FUNCTION_BLOCK CASE_SEQUENCER (* Solvability control: ecc_persistent form, designed by hand. Never shown to a model. *)
  (* Standard: 61499-2 *)
  (* Version 1.0, 2026-11-06, st2fb *)
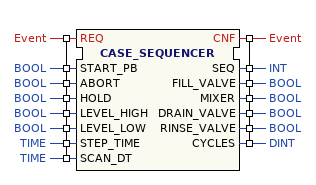
  EVENT_INPUT
    REQ WITH START_PB, ABORT, HOLD, LEVEL_HIGH, LEVEL_LOW, STEP_TIME, SCAN_DT;
  END_EVENT
  EVENT_OUTPUT
    CNF WITH SEQ, FILL_VALVE, MIXER, DRAIN_VALVE, RINSE_VALVE, CYCLES;
  END_EVENT
  VAR_INPUT
    START_PB : BOOL;
    ABORT : BOOL;
    HOLD : BOOL;
    LEVEL_HIGH : BOOL;
    LEVEL_LOW : BOOL;
    STEP_TIME : TIME;
    SCAN_DT : TIME;
  END_VAR
  VAR_OUTPUT
    SEQ : INT;
    FILL_VALVE : BOOL;
    MIXER : BOOL;
    DRAIN_VALVE : BOOL;
    RINSE_VALVE : BOOL;
    CYCLES : DINT;
  END_VAR
  VAR
    TIMING : BOOL;
    ST2FB_NOW : TIME;
    STEP_TIMER_IN : BOOL;
    STEP_TIMER_PT : TIME;
    STEP_TIMER_Q : BOOL;
    STEP_TIMER_ET : TIME;
    STEP_TIMER_STATE : INT;
    STEP_TIMER_PREV_IN : BOOL;
    STEP_TIMER_START_TIME : TIME;
  END_VAR
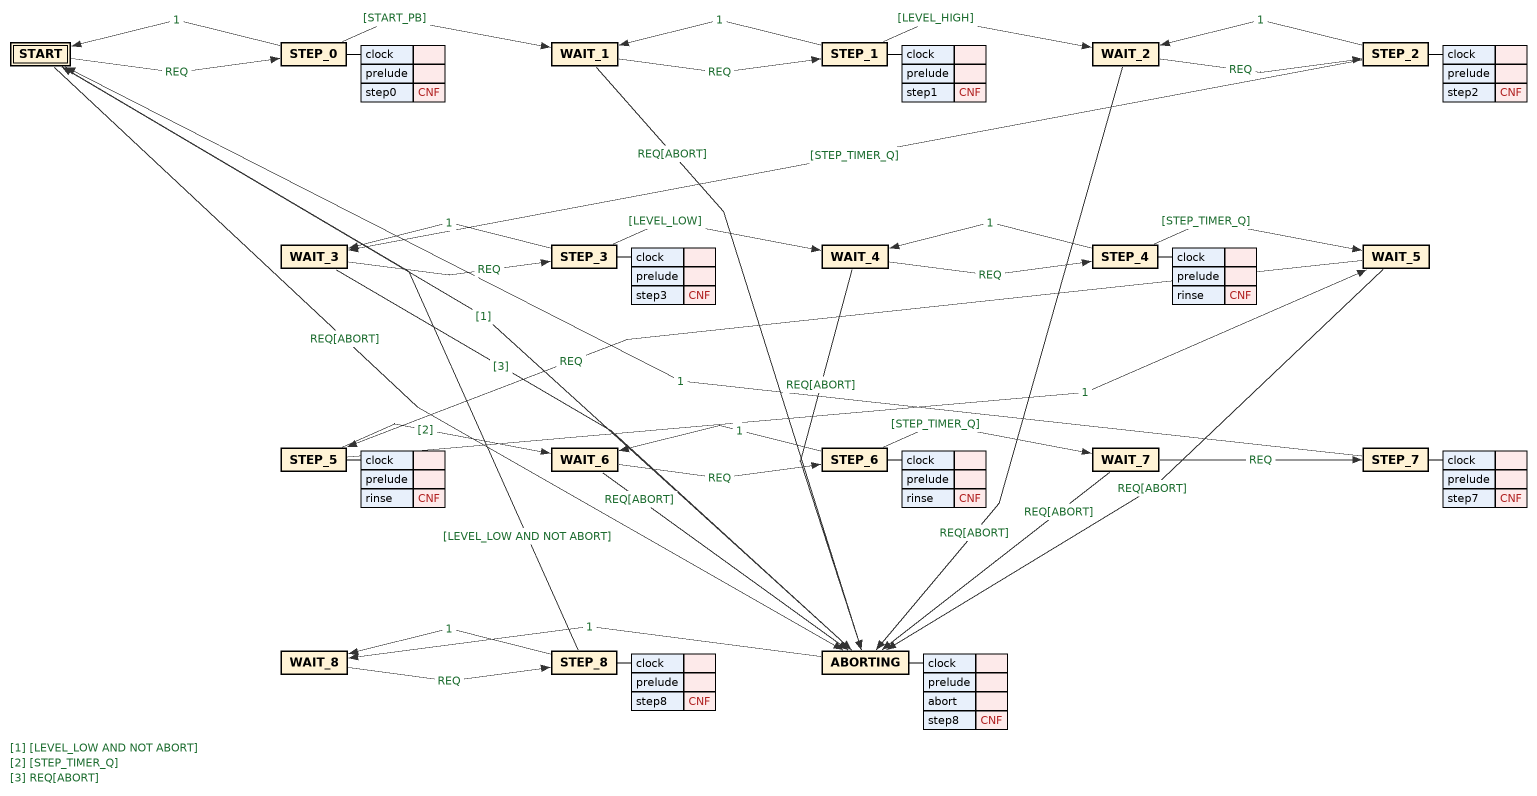
  EC_STATES
    START;
    STEP_0 : clock, prelude, step0 -> CNF;
    WAIT_1;
    STEP_1 : clock, prelude, step1 -> CNF;
    WAIT_2;
    STEP_2 : clock, prelude, step2 -> CNF;
    WAIT_3;
    STEP_3 : clock, prelude, step3 -> CNF;
    WAIT_4;
    STEP_4 : clock, prelude, rinse -> CNF;
    WAIT_5;
    STEP_5 : clock, prelude, rinse -> CNF;
    WAIT_6;
    STEP_6 : clock, prelude, rinse -> CNF;
    WAIT_7;
    STEP_7 : clock, prelude, step7 -> CNF;
    WAIT_8;
    STEP_8 : clock, prelude, step8 -> CNF;
    ABORTING : clock, prelude, abort, step8 -> CNF;
  END_STATES
  EC_TRANSITIONS
    START TO ABORTING := REQ[ABORT];
    START TO STEP_0 := REQ;
    WAIT_1 TO ABORTING := REQ[ABORT];
    WAIT_1 TO STEP_1 := REQ;
    WAIT_2 TO ABORTING := REQ[ABORT];
    WAIT_2 TO STEP_2 := REQ;
    WAIT_3 TO ABORTING := REQ[ABORT];
    WAIT_3 TO STEP_3 := REQ;
    WAIT_4 TO ABORTING := REQ[ABORT];
    WAIT_4 TO STEP_4 := REQ;
    WAIT_5 TO ABORTING := REQ[ABORT];
    WAIT_5 TO STEP_5 := REQ;
    WAIT_6 TO ABORTING := REQ[ABORT];
    WAIT_6 TO STEP_6 := REQ;
    WAIT_7 TO ABORTING := REQ[ABORT];
    WAIT_7 TO STEP_7 := REQ;
    WAIT_8 TO STEP_8 := REQ;
    STEP_0 TO WAIT_1 := [START_PB];
    STEP_0 TO START := 1;
    STEP_1 TO WAIT_2 := [LEVEL_HIGH];
    STEP_1 TO WAIT_1 := 1;
    STEP_2 TO WAIT_3 := [STEP_TIMER_Q];
    STEP_2 TO WAIT_2 := 1;
    STEP_3 TO WAIT_4 := [LEVEL_LOW];
    STEP_3 TO WAIT_3 := 1;
    STEP_4 TO WAIT_5 := [STEP_TIMER_Q];
    STEP_4 TO WAIT_4 := 1;
    STEP_5 TO WAIT_6 := [STEP_TIMER_Q];
    STEP_5 TO WAIT_5 := 1;
    STEP_6 TO WAIT_7 := [STEP_TIMER_Q];
    STEP_6 TO WAIT_6 := 1;
    STEP_7 TO START := 1;
    STEP_8 TO START := [LEVEL_LOW AND NOT ABORT];
    STEP_8 TO WAIT_8 := 1;
    ABORTING TO START := [LEVEL_LOW AND NOT ABORT];
    ABORTING TO WAIT_8 := 1;
  END_TRANSITIONS
  ALGORITHM clock IN ST:
ST2FB_NOW := ST2FB_NOW + SCAN_DT;
  END_ALGORITHM
  ALGORITHM prelude IN ST:
IF NOT HOLD THEN
  STEP_TIMER_IN := TIMING;
  STEP_TIMER_PT := STEP_TIME;
  IF STEP_TIMER_STATE = 0 AND NOT STEP_TIMER_PREV_IN AND STEP_TIMER_IN THEN
    STEP_TIMER_STATE := 1;
    STEP_TIMER_Q := FALSE;
    STEP_TIMER_START_TIME := ST2FB_NOW;
  ELSE
    IF NOT STEP_TIMER_IN THEN
      STEP_TIMER_ET := T#0s;
      STEP_TIMER_Q := FALSE;
      STEP_TIMER_STATE := 0;
    ELSIF STEP_TIMER_STATE = 1 THEN
      IF STEP_TIMER_START_TIME + STEP_TIMER_PT <= ST2FB_NOW THEN
        STEP_TIMER_STATE := 2;
        STEP_TIMER_Q := TRUE;
        STEP_TIMER_ET := STEP_TIMER_PT;
      ELSE
        STEP_TIMER_ET := ST2FB_NOW - STEP_TIMER_START_TIME;
      END_IF;
    END_IF;
  END_IF;
  STEP_TIMER_PREV_IN := STEP_TIMER_IN;
END_IF;
FILL_VALVE := FALSE;
MIXER := FALSE;
DRAIN_VALVE := FALSE;
RINSE_VALVE := FALSE;
  END_ALGORITHM
  ALGORITHM step0 IN ST:
TIMING := FALSE;
IF START_PB THEN
  SEQ := 1;
END_IF;
  END_ALGORITHM
  ALGORITHM step1 IN ST:
FILL_VALVE := TRUE;
IF LEVEL_HIGH THEN
  SEQ := 2;
  TIMING := TRUE;
END_IF;
  END_ALGORITHM
  ALGORITHM step2 IN ST:
MIXER := TRUE;
IF STEP_TIMER_Q THEN
  SEQ := 3;
  TIMING := FALSE;
END_IF;
  END_ALGORITHM
  ALGORITHM step3 IN ST:
DRAIN_VALVE := TRUE;
IF LEVEL_LOW THEN
  SEQ := 4;
END_IF;
  END_ALGORITHM
  ALGORITHM rinse IN ST:
RINSE_VALVE := TRUE;
IF STEP_TIMER_Q THEN
  SEQ := SEQ + 1;
  TIMING := FALSE;
ELSE
  TIMING := TRUE;
END_IF;
  END_ALGORITHM
  ALGORITHM step7 IN ST:
CYCLES := CYCLES + 1;
SEQ := 0;
  END_ALGORITHM
  ALGORITHM abort IN ST:
SEQ := 8;
  END_ALGORITHM
  ALGORITHM step8 IN ST:
TIMING := FALSE;
DRAIN_VALVE := TRUE;
IF LEVEL_LOW AND NOT ABORT THEN
  SEQ := 0;
END_IF;
  END_ALGORITHM
END_FUNCTION_BLOCK
